SUBAPPLICATION ALR_GT_0 (* Prüft ob LREAL-Adapter Wert > 0 ist (AX-Adapter Ausgang) *)
  (* Standard: 61499-2 *)
  (* Version 1.0, 2026-10-15, franz, Meisterschulen am Ostbahnhof *)
  PACKAGE MyLib::sys;
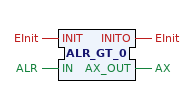
  EVENT_INPUT
    INIT : EInit; (* Initialization Request *)
  END_EVENT
  EVENT_OUTPUT
    INITO : EInit; (* Initialization Confirm *)
  END_EVENT
  SOCKETS
    IN : adapter::types::unidirectional::ALR;
  END_SOCKETS
  PLUGS
    AX_OUT : adapter::types::unidirectional::AX;
  END_PLUGS
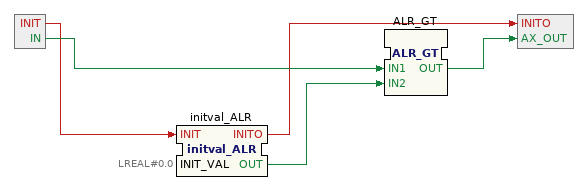
  FBS
    ALR_GT : adapter::iec61131::comparison::ALR_GT;
    initval_ALR : adapter::types::unidirectional::ALR::initval::initval_ALR(INIT_VAL := LREAL#0.0);
  END_FBS
  EVENT_CONNECTIONS
    INIT TO initval_ALR.INIT;
    initval_ALR.INITO TO INITO;
  END_CONNECTIONS
  ADAPTER_CONNECTIONS
    IN TO ALR_GT.IN1;
    ALR_GT.OUT TO AX_OUT;
    initval_ALR.OUT TO ALR_GT.IN2;
  END_CONNECTIONS
END_SUBAPPLICATION
